FUNCTION_BLOCK SimulatedActuator EXTENDS ActuatorBase
VAR
    _TravelTime   : TIME;
    _DrivenTarget : E_ActuatorTarget;
    _Travel       : TON;
    _IsStuck      : BOOL;
END_VAR
(*
    SimulatedActuator

    Stands in for a cylinder or gripper with end sensors. Reaches the
    commanded end TravelTime after the move starts. The supervision is
    ActuatorBase's, unchanged, so a move that never arrives faults exactly
    as a real one would. SetStuck() stops it moving. Has no I/O.
*)

METHOD FB_init : BOOL
VAR_INPUT
    bInitRetains : BOOL;
    bInCopyCode  : BOOL;
    Name         : STRING(32);
    MoveTimeout  : TIME;
    TravelTime   : TIME;
END_VAR
_TravelTime := TravelTime;
Configure(Name := Name, MoveTimeout := MoveTimeout);
END_METHOD

METHOD PUBLIC SetStuck
VAR_INPUT
    IsStuck : BOOL;
END_VAR
_IsStuck := IsStuck;
END_METHOD

METHOD PROTECTED IsWired : BOOL
IsWired := TRUE;                                    // nothing to wire
END_METHOD

METHOD PROTECTED DriveOutputs
VAR_INPUT
    Target : E_ActuatorTarget;
END_VAR
IF Target <> _DrivenTarget THEN
    _DrivenTarget := Target;
    _Travel(IN := FALSE);                           // a new move starts from the beginning
END_IF
_Travel(IN := Target <> E_ActuatorTarget.None AND NOT _IsStuck, PT := _TravelTime);
END_METHOD

METHOD PROTECTED IsAtPosition : BOOL
VAR_INPUT
    Position : E_ActuatorTarget;
END_VAR
IsAtPosition := Position <> E_ActuatorTarget.None AND Position = _DrivenTarget AND _Travel.Q;
END_METHOD

METHOD PROTECTED DriveSafe
_Travel(IN := FALSE);
END_METHOD

END_FUNCTION_BLOCK

(* stored: Version 1.1.0.1, ProductVersion 3.1.4026.0
   POU SimulatedActuator: Id {ac7c9dc8-0fef-4577-a3cc-72bd5e49513a}, SpecialFunc None
   Method FB_init: Id {5fa20193-0913-4b76-9672-a3f4cb9718cc}
   Method SetStuck: Id {95b7ad40-d702-4b8a-b1cc-5248ef6ca77d}
   Method IsWired: Id {71d07e8f-3473-488d-87b8-4b178dfb99e3}
   Method DriveOutputs: Id {526cc409-5a8d-4f42-b10c-1b9a4b9ff44f}
   Method IsAtPosition: Id {502484e1-d81a-4713-8a51-3f810359a5ee}
   Method DriveSafe: Id {ffbc2ddf-9b3f-4e61-96aa-cf632c6edc87} *)
